// TIA Portal V21 export
// export: Created 2026-11-10T19:16:53.147361Z, ExportSetting WithDefaults, DisplayName Totally Integrated Automation Portal, DisplayVersion V21 Update 3, DisplayName STEP 7 Professional, DisplayVersion V21 Update 3, DisplayName STEP 7 Safety, DisplayVersion V21, DisplayName Tech WebApplication, DisplayVersion V21, DisplayName WinCC Basic/Comfort/Advanced, DisplayVersion V21 Update 3, DisplayName WinCC Unified, DisplayVersion V21 Update 3
TYPE "UDT_Outer"
// stored: IsFailsafeCompliant false
   STRUCT
      inner { S7_SetPoint := 'True'} : "UDT_Inner";
      innerArr { S7_SetPoint := 'True'} : Array[0..1] of "UDT_Inner";
      s : Struct
         "a" : Bool;
         "m" : Array[0..1, 0..1] of Byte;
      END_STRUCT;
      txt : String[20] := 'outer';
   END_STRUCT;
END_TYPE
